// TIA Portal V21 export
// export: Created 2026-11-10T23:32:29.7994667Z, ExportSetting WithDefaults, DisplayName Totally Integrated Automation Portal, DisplayVersion V21 Update 3, DisplayName STEP 7 Professional, DisplayVersion V21 Update 3, DisplayName STEP 7 Safety, DisplayVersion V21, DisplayName Tech WebApplication, DisplayVersion V21, DisplayName WinCC Basic/Comfort/Advanced, DisplayVersion V21 Update 3, DisplayName WinCC Unified, DisplayVersion V21 Update 3
DATA_BLOCK "mTO_Interpreter"   // DB9, Motion_DB
// stored: AutoNumber true, DBAccessibleFromOPCUA true, DBAccessibleFromWebserver true, InstanceOfName TO_Interpreter, OfSystemLibElement TO_Interpreter, OfSystemLibVersion 8.0
TO_Interpreter   // technology object, version 8.0
   // // inherited from TO_Object
   // VAR
   //    ProgramName { ExternalWritable := 'False'} : Array[1..64] of DWord;
   //    MappingName { ExternalWritable := 'False'} : Array[1..64] of DWord;
   //    ProgramSource { ExternalWritable := 'False'} : DInt;
   //    MappingSource { ExternalWritable := 'False'} : DInt;
   //    ActualLineNumber { ExternalWritable := 'False'} : UDInt;
   //    Parameter { S7_SetPoint := 'True'} : TO_Struct_Interpreter_Parameter;
   //    Clipboard { S7_SetPoint := 'True'} : TO_Struct_Interpreter_Clipboard;
   //    StatusInterpreter { ExternalWritable := 'False'; S7_SetPoint := 'True'} : TO_Struct_Interpreter_StatusInterpreter;
   //    StatusWord { ExternalWritable := 'False'} : DWord;
   //    ErrorWord { ExternalWritable := 'False'} : DWord;
   //    ErrorDetail { ExternalWritable := 'False'; S7_SetPoint := 'True'} : TO_Struct_Interpreter_ErrorDetail;
   //    WarningWord { ExternalWritable := 'False'} : DWord;
   //    ControlPanel { S7_SetPoint := 'True'} : TO_Struct_Interpreter_ControlPanel;
   //    InternalToTrace { S7_SetPoint := 'True'} : Array[1..4] of TO_Struct_Internal;
   // END_VAR
BEGIN
END_DATA_BLOCK
